Fanuc KAREL source: kb00128.KL

PROGRAM KB00128
%STACKSIZE=65535
%PRIORITY=65535
%NOLOCKGROUP
VAR
P1 : POSITION
RESULT : VECTOR
BEGIN
RESULT=ORIENT(P1)
END KB00128
